// TwinCAT 3 PLC project AdsReadDemoPlc
// ProgramVersion: 3.1.4026.22
// libraries:
//   Tc2_Standard, * (Beckhoff Automation GmbH)
//   Tc2_System, * (Beckhoff Automation GmbH)
// project tree:
//   DUTs/ ST_Trigger.TcDUT
//   GVLs/ GVL_Param.TcGVL
//   POUs/ MAIN.TcPOU
//   / PlcTask.TcTTO
// real-time tasks:
//   TASK PlcTask: cycle T#10ms, priority 20, ADS port 350

CONFIGURATION AdsReadDemoPlc
    RESOURCE PLC ON TwinCAT3
        TASK PlcTask(INTERVAL := T#10ms, PRIORITY := 20);
        PROGRAM MAIN WITH PlcTask : MAIN;
    END_RESOURCE
END_CONFIGURATION

// ---- DUTs/ST_Trigger.TcDUT
// 模式 C / D 看的觸發值；兩個欄位同一個 cycle 寫入，C# 一次讀 12 bytes
{attribute 'pack_mode' := '1'}
TYPE ST_Trigger :
STRUCT
	nTrigger : UDINT; // 改值次數，每次 +1
	nPlcTime : ULINT; // 改值當下的 F_GetSystemTime() (100 ns, since 1601-01-01 UTC)
END_STRUCT
END_TYPE

// ---- GVLs/GVL_Param.TcGVL
{attribute 'qualified_only'}
VAR_GLOBAL CONSTANT
	cValueCount      : INT := 1000;                // MAIN.aValues 元素數 (模式 A / B 讀的量)
	cPhaseStepRad    : LREAL := 0.05;              // 每 cycle 相位增量 (rad)
	cElementPhaseRad : LREAL := 0.01;              // 相鄰元素的相位差 (rad)
	cTwoPiRad        : LREAL := 6.283185307179586; // 2π (rad)
	cTriggerPeriod   : TIME := T#2S;               // nTrigger 自動 +1 的預設間隔
END_VAR

// ---- POUs/MAIN.TcPOU
// ADS 讀變數示範的資料來源：aValues 每 cycle 更新 (模式 A / B)，stTrigger 定時或依 C# 要求 +1 (模式 C / D)
PROGRAM MAIN
VAR
	aValues          : ARRAY[1..GVL_Param.cValueCount] OF LREAL; // aValues[i] = i + SIN(相位)，每 cycle 都變
	stTrigger        : ST_Trigger;                               // 模式 C / D 讀這個 (12 bytes)
	bAutoTrigger     : BOOL := TRUE;                             // TRUE = 每 tTriggerPeriod 自動 +1；C# --trigger host 會改 FALSE
	tTriggerPeriod   : TIME := GVL_Param.cTriggerPeriod;         // 自動 +1 間隔，可從 ADS 改
	nHostRequest     : UDINT;                                    // C# --trigger host 寫入新值，下一個 cycle nTrigger +1
	nPlcTimeNow      : ULINT;                                    // 每 cycle 的 F_GetSystemTime() (100 ns)，C# 估時鐘差用
	nCycleCount      : UDINT;                                    // 本程式執行次數，看 task 是否真的在跑
	fPhaseRad        : LREAL;                                    // 目前相位 (rad), 0 ~ 2π
	fbTriggerTimer   : TON;
	nLastHostRequest : UDINT;
	bBump            : BOOL;
	nIndex           : INT;
END_VAR

nPlcTimeNow := F_GetSystemTime();
nCycleCount := nCycleCount + 1;

// 模式 A / B：1000 個 LREAL 每 cycle 都變，C# 讀到的值會不一樣
fPhaseRad := fPhaseRad + GVL_Param.cPhaseStepRad;
IF fPhaseRad >= GVL_Param.cTwoPiRad THEN
	fPhaseRad := fPhaseRad - GVL_Param.cTwoPiRad;
END_IF
FOR nIndex := 1 TO GVL_Param.cValueCount DO
	aValues[nIndex] := INT_TO_LREAL(nIndex) + SIN(fPhaseRad + INT_TO_LREAL(nIndex) * GVL_Param.cElementPhaseRad);
END_FOR

// 模式 C / D：定時 +1，或 C# 改了 nHostRequest 就 +1
fbTriggerTimer(IN := bAutoTrigger, PT := tTriggerPeriod);
bBump := fbTriggerTimer.Q;
IF fbTriggerTimer.Q THEN
	fbTriggerTimer(IN := FALSE); // 重新起算，下個 cycle 再開始計時
END_IF
IF nHostRequest <> nLastHostRequest THEN
	nLastHostRequest := nHostRequest;
	bBump := TRUE;
END_IF
IF bBump THEN
	stTrigger.nTrigger := stTrigger.nTrigger + 1;
	stTrigger.nPlcTime := nPlcTimeNow;
END_IF

END_PROGRAM
